Staubli VAL3: pointItem.dtx

public pointRx pPointRx[2]
  [0] = {fatherId=world[0]}
  [1] = {fatherId=world[0]}
public jointRx jJointRx
public paraItem pParaItem
  [0]
    mdesc mMdesc
    num nMoveType
    num nActionIndex
    num nPercentage
    ifItem iIfItem
      [0]
        num nSigType[3]
        num nSigIndex[3]
        num nValue[3]
        bool bANDOR[2]
    num nDelay
    num nSigValue
    bool bSafePoint
public string sID
public bool bMarked
public pointRx pInter = {fatherId=world[0]}
